// TIA Portal V21 export
// export: Created 2026-11-10T19:39:25.8680175Z, ExportSetting WithDefaults, DisplayName Totally Integrated Automation Portal, DisplayVersion V21 Update 3, DisplayName STEP 7 Professional, DisplayVersion V21 Update 3, DisplayName STEP 7 Safety, DisplayVersion V21, DisplayName Tech WebApplication, DisplayVersion V21, DisplayName WinCC Basic/Comfort/Advanced, DisplayVersion V21 Update 3, DisplayName WinCC Unified, DisplayVersion V21 Update 3
DATA_BLOCK "Motor1_DB"   // DB1
VERSION : 0.1
// stored: AutoNumber true, DBAccessibleFromOPCUA true, DBAccessibleFromWebserver true, InstanceOfName FB_Motor, InstanceOfType FB
"FB_Motor"
   // VAR_INPUT
   //    start : Bool;
   //    setSpeed : Real;
   // END_VAR
   // VAR_OUTPUT
   //    running : Bool;
   // END_VAR
   // VAR
   //    tOn { S7_SetPoint := 'True'} : TON_TIME;
   //    hours : DInt := 5;
   // END_VAR
BEGIN
END_DATA_BLOCK
